(* Provider test double that exposes the queue of ended spans for assertions. *)
FUNCTION_BLOCK FB_TracerProvider_ForInspection EXTENDS FB_TracerProvider

PROPERTY spans : REFERENCE TO FB_SpanQueue
GET
spans REF= THIS^._spans;
END_GET
END_PROPERTY

END_FUNCTION_BLOCK

(* stored: Version 1.1.0.1
   POU FB_TracerProvider_ForInspection: Id {64e232fc-bd17-42ef-92ba-3f806a11e717}, SpecialFunc None
   Property spans: Id {63e5096e-8ae5-44e1-a146-fa4f821b1b01}
   Get Get: Id {2d64f5ed-f657-4729-8a80-d9896532b8d8} *)
